Fanuc KAREL source: KT00622.KL

PROGRAM KT00622
%NOLOCKGROUP
VAR
  B1: BOOLEAN
  B2: BOOLEAN
  OUT: INTEGER
BEGIN
  B1 = TRUE
  B2 = FALSE
  B1 = TRUE
  B2 = FALSE
  OUT = - B1
END KT00622
